Fanuc TP program (LS listing): MAIN_1.LS

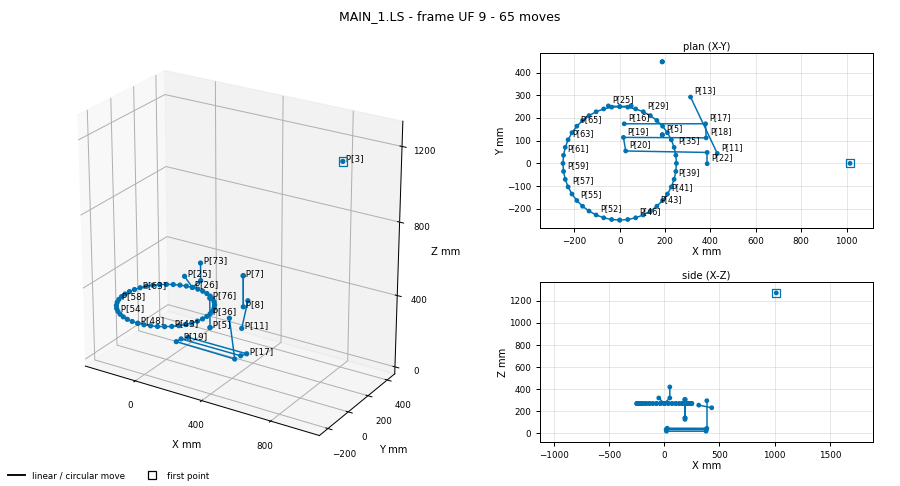
[picture p0: tool path of MAIN_1.LS in frame UF 9, 65 of 75 moves have a stored position in this frame; points joined in program order, loops and branches not executed]
/PROG  MAIN_1
/ATTR
OWNER		= MNEDITOR;
COMMENT		= "RoboDK sequence";
PROG_SIZE	= 0;
CREATE		= DATE 31-12-14  TIME 12:00:00;
MODIFIED	= DATE 31-12-14  TIME 12:00:00;
FILE_NAME	= MAIN_1;
VERSION		= 0;
LINE_COUNT	= 166;
MEMORY_SIZE	= 0;
PROTECT		= READ_WRITE;
TCD:  STACK_SIZE	= 0,
      TASK_PRIORITY	= 50,
      TIME_SLICE	= 0,
      BUSY_LAMP_OFF	= 0,
      ABORT_REQUEST	= 0,
      PAUSE_REQUEST	= 0;
DEFAULT_GROUP	= 1,*,*,*,*,*,*;
CONTROL_CODE	= 00000000 00000000;
/MN
   1:  ! Program generated by RoboDK v5.6.9 for RoboDK Industrial on 2 ;
   2:  ! 6/02/2024 09:58:20 ;
   3:  ! Using nominal kinematics. ;
   4:J P[1] 20% FINE ;
   5:J P[2] 20% FINE ;
   6:L P[3] 200mm/sec FINE ;
   7:  DO[5]=ON ;
   8:  DO[5]=ON ;
   9:  DO[5]=(0.5) ;
  10:  DO[5]=(true) ;
  11:  AO[5]=(1) ;
  12:  AO[5]=(2) ;
  13:  AO[5]=(0.5) ;
  14:  AO[5]=(true) ;
  15:  var=(val) ;
  16:  var=(val) ;
  17:  WAIT DI[5]=ON ;
  18:  WAIT DI[5]=ON ;
  19:  WAIT DI[5]=(0.5) ;
  20:  WAIT DI[5]=(true) ;
  21:  $WAITTMOUT=100 ;
  22:  WAIT DI[5]=ON TIMEOUT, LBL[1] ;
  23:  MESSAGE[Timed out for LBL 1] ;
  24:  PAUSE ;
  25:  LBL[1] ;
  26:  WAIT var=(val) ;
  27:  $WAITTMOUT=100 ;
  28:  WAIT var=(val) TIMEOUT, LBL[2] ;
  29:  MESSAGE[Timed out for LBL 2] ;
  30:  PAUSE ;
  31:  LBL[2] ;
  32:  MESSAGE[Message] ;
  33:  CALL REMOTE_PROG_ ;
  34:  CODE_INSERT_172;
  35:  ! Insert Comment ;
  36:  PR[9,1]=719.013 ;
  37:  PR[9,2]=-664.003 ;
  38:  PR[9,3]=0.000 ;
  39:  PR[9,4]=0.000 ;
  40:  PR[9,5]=0.000 ;
  41:  PR[9,6]=0.000 ;
  42:  UFRAME[9]=PR[9] ;
  43:  UFRAME_NUM=9 ;
  44:  UTOOL_NUM=1 ;
  45:  ! UT1:129.1,0.0,85.5,0.0,22.8,0.0 ;
  46:J P[4] 100% CNT10 ACC100 ;
  47:L P[5] 100mm/sec FINE ACC100 ;
  48:  DO[5]=ON ;
  49:  CALL PICK_PART_11 ;
  50:L P[6] 300mm/sec CNT10 ACC100 ;
  51:L P[7] 300mm/sec CNT10 ACC100 ;
  52:  ! MoveSearch command not implemented ;
  53:L P[8] 100mm/sec FINE ACC100 ;
  54:  DO[5]=OFF ;
  55:  CALL PLACE_PART_1 ;
  56:L P[9] 100mm/sec CNT10 ACC100 ;
  57:  PR[9,1]=577.670 ;
  58:  PR[9,2]=392.250 ;
  59:  PR[9,3]=0.000 ;
  60:  PR[9,4]=0.000 ;
  61:  PR[9,5]=0.000 ;
  62:  PR[9,6]=38.960 ;
  63:  UFRAME[9]=PR[9] ;
  64:  UFRAME_NUM=9 ;
  65:J P[10] 2% CNT25 ACC100 ;
  66:C P[11]
       P[12] 100mm/sec CNT25 ;
  67:  ! Circular movement using joint targets is not supported. Chang ;
  68:  ! e the target type to cartesian or use a joint movement. ;
  69:L P[13] 100mm/sec FINE ACC100 ;
  70:J P[14] 2% FINE ACC100 ;
  71:  PR[9,1]=0.000 ;
  72:  PR[9,2]=782.714 ;
  73:  PR[9,3]=377.610 ;
  74:  PR[9,4]=0.000 ;
  75:  PR[9,5]=0.000 ;
  76:  PR[9,6]=0.000 ;
  77:  UFRAME[9]=PR[9] ;
  78:  UFRAME_NUM=9 ;
  79:J P[15] 2% FINE ACC100 ;
  80:L P[16] 100mm/sec FINE ACC100 ;
  81:L P[17] 100mm/sec FINE ACC100 ;
  82:L P[18] 100mm/sec FINE ACC100 ;
  83:L P[19] 100mm/sec FINE ACC100 ;
  84:L P[20] 100mm/sec FINE ACC100 ;
  85:L P[21] 100mm/sec FINE ACC100 ;
  86:L P[22] 100mm/sec FINE ACC100 ;
  87:J P[23] 2% FINE ACC100 ;
  88:  CALL EVENT_PROG_S ;
  89:  PR[9,1]=13.637 ;
  90:  PR[9,2]=-840.080 ;
  91:  PR[9,3]=0.000 ;
  92:  PR[9,4]=0.000 ;
  93:  PR[9,5]=0.000 ;
  94:  PR[9,6]=-90.000 ;
  95:  UFRAME[9]=PR[9] ;
  96:  UFRAME_NUM=9 ;
  97:  ! Show Tool 1 ;
  98:J P[24] 20% FINE ACC100 ;
  99:  CALL EVENT_PATH_A ;
 100:L P[25] 1000mm/sec CNT1 ACC100 ;
 101:L P[26] 1000mm/sec FINE ACC100 ;
 102:  CALL EVENT_PATH_S ;
 103:L P[27] 50mm/sec CNT1 ACC100 ;
 104:L P[28] 50mm/sec CNT1 ACC100 ;
 105:L P[29] 50mm/sec CNT1 ACC100 ;
 106:L P[30] 50mm/sec CNT1 ACC100 ;
 107:L P[31] 50mm/sec CNT1 ACC100 ;
 108:L P[32] 50mm/sec CNT1 ACC100 ;
 109:L P[33] 50mm/sec CNT1 ACC100 ;
 110:L P[34] 50mm/sec CNT1 ACC100 ;
 111:L P[35] 50mm/sec CNT1 ACC100 ;
 112:L P[36] 50mm/sec CNT1 ACC100 ;
 113:L P[37] 50mm/sec CNT1 ACC100 ;
 114:L P[38] 50mm/sec CNT1 ACC100 ;
 115:L P[39] 50mm/sec CNT1 ACC100 ;
 116:L P[40] 50mm/sec CNT1 ACC100 ;
 117:L P[41] 50mm/sec CNT1 ACC100 ;
 118:L P[42] 50mm/sec CNT1 ACC100 ;
 119:L P[43] 50mm/sec CNT1 ACC100 ;
 120:L P[44] 50mm/sec CNT1 ACC100 ;
 121:L P[45] 50mm/sec CNT1 ACC100 ;
 122:L P[46] 50mm/sec CNT1 ACC100 ;
 123:L P[47] 50mm/sec CNT1 ACC100 ;
 124:L P[48] 50mm/sec CNT1 ACC100 ;
 125:L P[49] 50mm/sec CNT1 ACC100 ;
 126:L P[50] 50mm/sec CNT1 ACC100 ;
 127:L P[51] 50mm/sec CNT1 ACC100 ;
 128:L P[52] 50mm/sec CNT1 ACC100 ;
 129:L P[53] 50mm/sec CNT1 ACC100 ;
 130:L P[54] 50mm/sec CNT1 ACC100 ;
 131:L P[55] 50mm/sec CNT1 ACC100 ;
 132:L P[56] 50mm/sec CNT1 ACC100 ;
 133:L P[57] 50mm/sec CNT1 ACC100 ;
 134:L P[58] 50mm/sec CNT1 ACC100 ;
 135:L P[59] 50mm/sec CNT1 ACC100 ;
 136:L P[60] 50mm/sec CNT1 ACC100 ;
 137:L P[61] 50mm/sec CNT1 ACC100 ;
 138:L P[62] 50mm/sec CNT1 ACC100 ;
 139:L P[63] 50mm/sec CNT1 ACC100 ;
 140:L P[64] 50mm/sec CNT1 ACC100 ;
 141:L P[65] 50mm/sec CNT1 ACC100 ;
 142:L P[66] 50mm/sec CNT1 ACC100 ;
 143:L P[67] 50mm/sec CNT1 ACC100 ;
 144:L P[68] 50mm/sec CNT1 ACC100 ;
 145:L P[69] 50mm/sec CNT1 ACC100 ;
 146:L P[70] 50mm/sec CNT1 ACC100 ;
 147:L P[71] 50mm/sec FINE ACC100 ;
 148:  CALL EVENT_PATH_F ;
 149:L P[72] 1000mm/sec CNT1 ACC100 ;
 150:L P[73] 1000mm/sec FINE ACC100 ;
 151:  CALL EVENT_PATH_R ;
 152:  CALL EVENT_PROG_F ;
 153:  PR[9,1]=719.013 ;
 154:  PR[9,2]=-664.003 ;
 155:  PR[9,3]=0.000 ;
 156:  PR[9,4]=0.000 ;
 157:  PR[9,5]=0.000 ;
 158:  PR[9,6]=0.000 ;
 159:  UFRAME[9]=PR[9] ;
 160:  UFRAME_NUM=9 ;
 161:J P[74] 20% CNT1 ACC100 ;
 162:  WAIT  1.25(sec) ;
 163:L P[75] 1000mm/sec CNT1 ACC100 ;
 164:  WAIT DI[1]=ON ;
 165:L P[76] 1000mm/sec FINE ACC100 ;
 166:  CALL PROG1_withav ;
/POS
P[1]{
   GP1:
    UF : 9, UT : 9,
	J1=    -0.000 deg,	J2=    0.000 deg,	J3=    0.000 deg,
	J4=    0.000 deg,	J5=    0.000 deg,	J6=    -0.000 deg
};
P[2]{
   GP1:
    UF : 9, UT : 9,
	J1=    0.000 deg,	J2=    3.211 deg,	J3=    -15.424 deg,
	J4=    0.000 deg,	J5=    12.213 deg,	J6=    -0.000 deg
};
P[3]{
   GP1:
    UF : 9, UT : 9,        CONFIG : 'F U T, 0, 0, 0',
	X =  1015.000  mm,	Y =     0.000  mm,	Z =  1272.000  mm,
	W =     0.000 deg,	P =    90.000 deg,	R =     0.000 deg
};
P[4]{
   GP1:
    UF : 9, UT : 1,
	J1=    -29.332 deg,	J2=    46.677 deg,	J3=    -0.025 deg,
	J4=    26.546 deg,	J5=    25.396 deg,	J6=    -51.634 deg
};
P[5]{
   GP1:
    UF : 9, UT : 1,        CONFIG : 'N U T, 0, 0, 0',
	X =   187.786  mm,	Y =   125.499  mm,	Z =   139.112  mm,
	W =   179.996 deg,	P =     0.180 deg,	R =  -179.997 deg
};
P[6]{
   GP1:
    UF : 9, UT : 1,
	J1=    -29.332 deg,	J2=    46.677 deg,	J3=    -0.024 deg,
	J4=    26.546 deg,	J5=    25.396 deg,	J6=    -51.634 deg
};
P[7]{
   GP1:
    UF : 9, UT : 1,        CONFIG : 'N U T, 0, 0, 0',
	X =   187.272  mm,	Y =   447.522  mm,	Z =   305.347  mm,
	W =  -179.998 deg,	P =     0.185 deg,	R =   179.999 deg
};
P[8]{
   GP1:
    UF : 9, UT : 1,        CONFIG : 'N U T, 0, 0, 0',
	X =   187.851  mm,	Y =   447.517  mm,	Z =   126.235  mm,
	W =  -179.998 deg,	P =     0.185 deg,	R =   179.999 deg
};
P[9]{
   GP1:
    UF : 9, UT : 1,        CONFIG : 'N U T, 0, 0, 0',
	X =   187.272  mm,	Y =   447.522  mm,	Z =   305.347  mm,
	W =  -179.998 deg,	P =     0.185 deg,	R =   179.999 deg
};
P[10]{
   GP1:
    UF : 9, UT : 1,
	J1=    52.186 deg,	J2=    45.676 deg,	J3=    6.920 deg,
	J4=    66.734 deg,	J5=    19.932 deg,	J6=    -92.730 deg
};
P[11]{
   GP1:
    UF : 9, UT : 1,        CONFIG : 'N U T, 0, 0, 0',
	X =   430.047  mm,	Y =    43.774  mm,	Z =   231.503  mm,
	W =   178.913 deg,	P =    11.181 deg,	R =  -134.549 deg
};
P[12]{
   GP1:
    UF : 9, UT : 1,        CONFIG : 'N U T, 0, 0, 0',
	X =   109.688  mm,	Y =  -153.222  mm,	Z =   161.073  mm,
	W =   178.913 deg,	P =    11.181 deg,	R =  -134.549 deg
};
P[13]{
   GP1:
    UF : 9, UT : 1,        CONFIG : 'N U T, 0, 0, 0',
	X =   312.208  mm,	Y =   292.214  mm,	Z =   255.156  mm,
	W =   178.913 deg,	P =    11.181 deg,	R =  -134.549 deg
};
P[14]{
   GP1:
    UF : 9, UT : 1,
	J1=    -0.000 deg,	J2=    0.000 deg,	J3=    0.000 deg,
	J4=    0.000 deg,	J5=    0.000 deg,	J6=    -0.000 deg
};
P[15]{
   GP1:
    UF : 9, UT : 1,
	J1=    88.676 deg,	J2=    29.602 deg,	J3=    -6.429 deg,
	J4=    -1.984 deg,	J5=    49.479 deg,	J6=    4.548 deg
};
P[16]{
   GP1:
    UF : 9, UT : 1,        CONFIG : 'N U T, 0, 0, 0',
	X =    19.898  mm,	Y =   174.307  mm,	Z =    19.008  mm,
	W =  -179.533 deg,	P =    -5.426 deg,	R =   -94.928 deg
};
P[17]{
   GP1:
    UF : 9, UT : 1,        CONFIG : 'N U T, 0, 0, 0',
	X =   378.402  mm,	Y =   174.416  mm,	Z =    18.997  mm,
	W =  -179.533 deg,	P =    -5.426 deg,	R =   -94.928 deg
};
P[18]{
   GP1:
    UF : 9, UT : 1,        CONFIG : 'N U T, 0, 0, 0',
	X =   380.996  mm,	Y =   112.363  mm,	Z =    34.882  mm,
	W =  -178.348 deg,	P =   -18.136 deg,	R =   -95.294 deg
};
P[19]{
   GP1:
    UF : 9, UT : 1,        CONFIG : 'N U T, 0, 0, 0',
	X =    16.551  mm,	Y =   114.359  mm,	Z =    34.226  mm,
	W =  -178.348 deg,	P =   -18.136 deg,	R =   -95.294 deg
};
P[20]{
   GP1:
    UF : 9, UT : 1,        CONFIG : 'N U T, 0, 0, 0',
	X =    26.434  mm,	Y =    54.524  mm,	Z =    46.072  mm,
	W =   179.585 deg,	P =     4.348 deg,	R =   -95.461 deg
};
P[21]{
   GP1:
    UF : 9, UT : 1,        CONFIG : 'N U T, 0, 0, 0',
	X =   385.448  mm,	Y =    48.050  mm,	Z =    45.137  mm,
	W =   178.913 deg,	P =    11.181 deg,	R =   -95.590 deg
};
P[22]{
   GP1:
    UF : 9, UT : 1,        CONFIG : 'N U T, 0, 0, 0',
	X =   385.448  mm,	Y =    -1.625  mm,	Z =   295.251  mm,
	W =   178.913 deg,	P =    11.181 deg,	R =   -95.590 deg
};
P[23]{
   GP1:
    UF : 9, UT : 1,
	J1=    -0.000 deg,	J2=    0.000 deg,	J3=    0.000 deg,
	J4=    0.000 deg,	J5=    0.000 deg,	J6=    -0.000 deg
};
P[24]{
   GP1:
    UF : 9, UT : 1,
	J1=    -68.090 deg,	J2=    24.202 deg,	J3=    26.785 deg,
	J4=    38.213 deg,	J5=    36.202 deg,	J6=    -98.796 deg
};
P[25]{
   GP1:
    UF : 9, UT : 1,        CONFIG : 'N U T, 0, 0, 0',
	X =   -49.895  mm,	Y =   253.259  mm,	Z =   319.999  mm,
	W =  -179.975 deg,	P =     0.353 deg,	R =   -90.000 deg
};
P[26]{
   GP1:
    UF : 9, UT : 1,        CONFIG : 'N U T, 0, 0, 0',
	X =     0.000  mm,	Y =   250.000  mm,	Z =   270.000  mm,
	W =  -179.975 deg,	P =     0.353 deg,	R =   -90.000 deg
};
P[27]{
   GP1:
    UF : 9, UT : 1,        CONFIG : 'N U T, 0, 0, 0',
	X =    35.579  mm,	Y =   247.455  mm,	Z =   270.000  mm,
	W =  -179.925 deg,	P =     0.345 deg,	R =   -90.000 deg
};
P[28]{
   GP1:
    UF : 9, UT : 1,        CONFIG : 'N U T, 0, 0, 0',
	X =    70.433  mm,	Y =   239.873  mm,	Z =   270.000  mm,
	W =  -179.876 deg,	P =     0.331 deg,	R =   -89.999 deg
};
P[29]{
   GP1:
    UF : 9, UT : 1,        CONFIG : 'N U T, 0, 0, 0',
	X =   103.854  mm,	Y =   227.408  mm,	Z =   270.000  mm,
	W =  -179.831 deg,	P =     0.310 deg,	R =   -89.999 deg
};
P[30]{
   GP1:
    UF : 9, UT : 1,        CONFIG : 'N U T, 0, 0, 0',
	X =   135.160  mm,	Y =   210.313  mm,	Z =   270.000  mm,
	W =  -179.788 deg,	P =     0.283 deg,	R =   -89.999 deg
};
P[31]{
   GP1:
    UF : 9, UT : 1,        CONFIG : 'N U T, 0, 0, 0',
	X =   163.715  mm,	Y =   188.937  mm,	Z =   270.000  mm,
	W =  -179.750 deg,	P =     0.250 deg,	R =   -89.999 deg
};
P[32]{
   GP1:
    UF : 9, UT : 1,        CONFIG : 'N U T, 0, 0, 0',
	X =   188.937  mm,	Y =   163.715  mm,	Z =   270.000  mm,
	W =  -179.717 deg,	P =     0.212 deg,	R =   -89.999 deg
};
P[33]{
   GP1:
    UF : 9, UT : 1,        CONFIG : 'N U T, 0, 0, 0',
	X =   210.313  mm,	Y =   135.160  mm,	Z =   270.000  mm,
	W =  -179.689 deg,	P =     0.170 deg,	R =   -89.999 deg
};
P[34]{
   GP1:
    UF : 9, UT : 1,        CONFIG : 'N U T, 0, 0, 0',
	X =   227.408  mm,	Y =   103.854  mm,	Z =   270.000  mm,
	W =  -179.668 deg,	P =     0.124 deg,	R =   -89.999 deg
};
P[35]{
   GP1:
    UF : 9, UT : 1,        CONFIG : 'N U T, 0, 0, 0',
	X =   239.873  mm,	Y =    70.433  mm,	Z =   270.000  mm,
	W =  -179.654 deg,	P =     0.075 deg,	R =   -90.000 deg
};
P[36]{
   GP1:
    UF : 9, UT : 1,        CONFIG : 'N U T, 0, 0, 0',
	X =   247.455  mm,	Y =    35.579  mm,	Z =   270.000  mm,
	W =  -179.647 deg,	P =     0.025 deg,	R =   -90.000 deg
};
P[37]{
   GP1:
    UF : 9, UT : 1,        CONFIG : 'N U T, 0, 0, 0',
	X =   250.000  mm,	Y =     0.000  mm,	Z =   270.000  mm,
	W =  -179.647 deg,	P =    -0.025 deg,	R =   -90.000 deg
};
P[38]{
   GP1:
    UF : 9, UT : 1,        CONFIG : 'N U T, 0, 0, 0',
	X =   247.455  mm,	Y =   -35.579  mm,	Z =   270.000  mm,
	W =  -179.654 deg,	P =    -0.075 deg,	R =   -90.000 deg
};
P[39]{
   GP1:
    UF : 9, UT : 1,        CONFIG : 'N U T, 0, 0, 0',
	X =   239.873  mm,	Y =   -70.433  mm,	Z =   270.000  mm,
	W =  -179.668 deg,	P =    -0.124 deg,	R =   -90.001 deg
};
P[40]{
   GP1:
    UF : 9, UT : 1,        CONFIG : 'N U T, 0, 0, 0',
	X =   227.408  mm,	Y =  -103.854  mm,	Z =   270.000  mm,
	W =  -179.689 deg,	P =    -0.170 deg,	R =   -90.001 deg
};
P[41]{
   GP1:
    UF : 9, UT : 1,        CONFIG : 'N U T, 0, 0, 0',
	X =   210.313  mm,	Y =  -135.160  mm,	Z =   270.000  mm,
	W =  -179.717 deg,	P =    -0.212 deg,	R =   -90.001 deg
};
P[42]{
   GP1:
    UF : 9, UT : 1,        CONFIG : 'N U T, 0, 0, 0',
	X =   188.937  mm,	Y =  -163.715  mm,	Z =   270.000  mm,
	W =  -179.750 deg,	P =    -0.250 deg,	R =   -90.001 deg
};
P[43]{
   GP1:
    UF : 9, UT : 1,        CONFIG : 'N U T, 0, 0, 0',
	X =   163.715  mm,	Y =  -188.937  mm,	Z =   270.000  mm,
	W =  -179.788 deg,	P =    -0.283 deg,	R =   -90.001 deg
};
P[44]{
   GP1:
    UF : 9, UT : 1,        CONFIG : 'N U T, 0, 0, 0',
	X =   135.160  mm,	Y =  -210.313  mm,	Z =   270.000  mm,
	W =  -179.830 deg,	P =    -0.311 deg,	R =   -90.001 deg
};
P[45]{
   GP1:
    UF : 9, UT : 1,        CONFIG : 'N U T, 0, 0, 0',
	X =   103.854  mm,	Y =  -227.408  mm,	Z =   270.000  mm,
	W =  -179.876 deg,	P =    -0.332 deg,	R =   -90.001 deg
};
P[46]{
   GP1:
    UF : 9, UT : 1,        CONFIG : 'N U T, 0, 0, 0',
	X =    70.433  mm,	Y =  -239.873  mm,	Z =   270.000  mm,
	W =  -179.925 deg,	P =    -0.346 deg,	R =   -90.000 deg
};
P[47]{
   GP1:
    UF : 9, UT : 1,        CONFIG : 'N U T, 0, 0, 0',
	X =    35.579  mm,	Y =  -247.455  mm,	Z =   270.000  mm,
	W =  -179.975 deg,	P =    -0.353 deg,	R =   -90.000 deg
};
P[48]{
   GP1:
    UF : 9, UT : 1,        CONFIG : 'N U T, 0, 0, 0',
	X =     0.000  mm,	Y =  -250.000  mm,	Z =   270.000  mm,
	W =  -179.975 deg,	P =    -0.353 deg,	R =   -90.000 deg
};
P[49]{
   GP1:
    UF : 9, UT : 1,        CONFIG : 'N U T, 0, 0, 0',
	X =     0.000  mm,	Y =  -250.000  mm,	Z =   270.000  mm,
	W =   179.975 deg,	P =    -0.353 deg,	R =   -90.000 deg
};
P[50]{
   GP1:
    UF : 9, UT : 1,        CONFIG : 'N U T, 0, 0, 0',
	X =   -35.579  mm,	Y =  -247.455  mm,	Z =   270.000  mm,
	W =   179.925 deg,	P =    -0.346 deg,	R =   -90.000 deg
};
P[51]{
   GP1:
    UF : 9, UT : 1,        CONFIG : 'N U T, 0, 0, 0',
	X =   -70.433  mm,	Y =  -239.873  mm,	Z =   270.000  mm,
	W =   179.876 deg,	P =    -0.331 deg,	R =   -89.999 deg
};
P[52]{
   GP1:
    UF : 9, UT : 1,        CONFIG : 'N U T, 0, 0, 0',
	X =  -103.854  mm,	Y =  -227.408  mm,	Z =   270.000  mm,
	W =   179.831 deg,	P =    -0.310 deg,	R =   -89.999 deg
};
P[53]{
   GP1:
    UF : 9, UT : 1,        CONFIG : 'N U T, 0, 0, 0',
	X =  -135.160  mm,	Y =  -210.313  mm,	Z =   270.000  mm,
	W =   179.788 deg,	P =    -0.283 deg,	R =   -89.999 deg
};
P[54]{
   GP1:
    UF : 9, UT : 1,        CONFIG : 'N U T, 0, 0, 0',
	X =  -163.715  mm,	Y =  -188.937  mm,	Z =   270.000  mm,
	W =   179.750 deg,	P =    -0.250 deg,	R =   -89.999 deg
};
P[55]{
   GP1:
    UF : 9, UT : 1,        CONFIG : 'N U T, 0, 0, 0',
	X =  -188.937  mm,	Y =  -163.715  mm,	Z =   270.000  mm,
	W =   179.717 deg,	P =    -0.212 deg,	R =   -89.999 deg
};
P[56]{
   GP1:
    UF : 9, UT : 1,        CONFIG : 'N U T, 0, 0, 0',
	X =  -210.313  mm,	Y =  -135.160  mm,	Z =   270.000  mm,
	W =   179.690 deg,	P =    -0.169 deg,	R =   -89.999 deg
};
P[57]{
   GP1:
    UF : 9, UT : 1,        CONFIG : 'N U T, 0, 0, 0',
	X =  -227.408  mm,	Y =  -103.854  mm,	Z =   270.000  mm,
	W =   179.669 deg,	P =    -0.123 deg,	R =   -89.999 deg
};
P[58]{
   GP1:
    UF : 9, UT : 1,        CONFIG : 'N U T, 0, 0, 0',
	X =  -239.873  mm,	Y =   -70.433  mm,	Z =   270.000  mm,
	W =   179.654 deg,	P =    -0.075 deg,	R =   -90.000 deg
};
P[59]{
   GP1:
    UF : 9, UT : 1,        CONFIG : 'N U T, 0, 0, 0',
	X =  -247.455  mm,	Y =   -35.579  mm,	Z =   270.000  mm,
	W =   179.647 deg,	P =    -0.025 deg,	R =   -90.000 deg
};
P[60]{
   GP1:
    UF : 9, UT : 1,        CONFIG : 'N U T, 0, 0, 0',
	X =  -250.000  mm,	Y =     0.000  mm,	Z =   270.000  mm,
	W =   179.647 deg,	P =     0.025 deg,	R =   -90.000 deg
};
P[61]{
   GP1:
    UF : 9, UT : 1,        CONFIG : 'N U T, 0, 0, 0',
	X =  -247.455  mm,	Y =    35.579  mm,	Z =   270.000  mm,
	W =   179.655 deg,	P =     0.075 deg,	R =   -90.000 deg
};
P[62]{
   GP1:
    UF : 9, UT : 1,        CONFIG : 'N U T, 0, 0, 0',
	X =  -239.873  mm,	Y =    70.433  mm,	Z =   270.000  mm,
	W =   179.669 deg,	P =     0.123 deg,	R =   -90.001 deg
};
P[63]{
   GP1:
    UF : 9, UT : 1,        CONFIG : 'N U T, 0, 0, 0',
	X =  -227.408  mm,	Y =   103.854  mm,	Z =   270.000  mm,
	W =   179.689 deg,	P =     0.170 deg,	R =   -90.001 deg
};
P[64]{
   GP1:
    UF : 9, UT : 1,        CONFIG : 'N U T, 0, 0, 0',
	X =  -210.313  mm,	Y =   135.160  mm,	Z =   270.000  mm,
	W =   179.717 deg,	P =     0.212 deg,	R =   -90.001 deg
};
P[65]{
   GP1:
    UF : 9, UT : 1,        CONFIG : 'N U T, 0, 0, 0',
	X =  -188.937  mm,	Y =   163.715  mm,	Z =   270.000  mm,
	W =   179.750 deg,	P =     0.250 deg,	R =   -90.001 deg
};
P[66]{
   GP1:
    UF : 9, UT : 1,        CONFIG : 'N U T, 0, 0, 0',
	X =  -163.715  mm,	Y =   188.937  mm,	Z =   270.000  mm,
	W =   179.788 deg,	P =     0.283 deg,	R =   -90.001 deg
};
P[67]{
   GP1:
    UF : 9, UT : 1,        CONFIG : 'N U T, 0, 0, 0',
	X =  -135.160  mm,	Y =   210.313  mm,	Z =   270.000  mm,
	W =   179.831 deg,	P =     0.310 deg,	R =   -90.001 deg
};
P[68]{
   GP1:
    UF : 9, UT : 1,        CONFIG : 'N U T, 0, 0, 0',
	X =  -103.854  mm,	Y =   227.408  mm,	Z =   270.000  mm,
	W =   179.876 deg,	P =     0.332 deg,	R =   -90.001 deg
};
P[69]{
   GP1:
    UF : 9, UT : 1,        CONFIG : 'N U T, 0, 0, 0',
	X =   -70.433  mm,	Y =   239.873  mm,	Z =   270.000  mm,
	W =   179.925 deg,	P =     0.346 deg,	R =   -90.000 deg
};
P[70]{
   GP1:
    UF : 9, UT : 1,        CONFIG : 'N U T, 0, 0, 0',
	X =   -35.579  mm,	Y =   247.455  mm,	Z =   270.000  mm,
	W =   179.975 deg,	P =     0.353 deg,	R =   -90.000 deg
};
P[71]{
   GP1:
    UF : 9, UT : 1,        CONFIG : 'N U T, 0, 0, 0',
	X =     0.000  mm,	Y =   250.000  mm,	Z =   270.000  mm,
	W =   179.975 deg,	P =     0.353 deg,	R =   -90.000 deg
};
P[72]{
   GP1:
    UF : 9, UT : 1,        CONFIG : 'N U T, 0, 0, 0',
	X =    49.895  mm,	Y =   253.258  mm,	Z =   319.999  mm,
	W =   179.975 deg,	P =     0.353 deg,	R =   -90.000 deg
};
P[73]{
   GP1:
    UF : 9, UT : 1,        CONFIG : 'N U T, 0, 0, 0',
	X =    49.939  mm,	Y =   252.642  mm,	Z =   419.997  mm,
	W =   179.975 deg,	P =     0.353 deg,	R =   -90.000 deg
};
P[74]{
   GP1:
    UF : 9, UT : 1,
	J1=    -29.332 deg,	J2=    46.677 deg,	J3=    -0.025 deg,
	J4=    26.546 deg,	J5=    25.396 deg,	J6=    -51.634 deg
};
P[75]{
   GP1:
    UF : 9, UT : 1,        CONFIG : 'N U T, 0, 0, 0',
	X =   187.786  mm,	Y =   125.499  mm,	Z =   139.112  mm,
	W =   179.996 deg,	P =     0.180 deg,	R =  -179.997 deg
};
P[76]{
   GP1:
    UF : 9, UT : 1,        CONFIG : 'N U T, 0, 0, 0',
	X =   187.264  mm,	Y =   125.487  mm,	Z =   305.356  mm,
	W =  -180.000 deg,	P =     0.184 deg,	R =   180.000 deg
};
/END
